// TIA Portal V15.1 export
// export: Created 2000-01-01T00:00:00.0000000Z, ExportSetting None
FUNCTION "FC_Rung" : Void   // FC42, LAD
{ S7_Optimized_Access := 'TRUE' }
   VAR_INPUT
      Local : Int;
   END_VAR
BEGIN

REGION Network 1
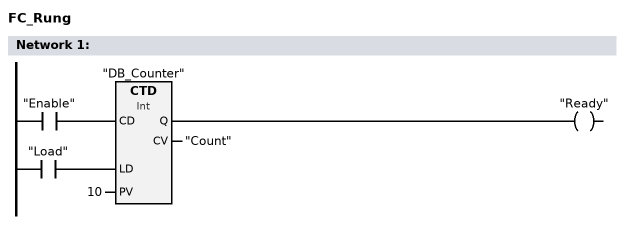
   RUNG wire#powerrail
      Contact( "Enable" )
      { S7_Templates := "value_type := Int" } "DB_Counter".CTD(ld := wire#w1, pv := 10, cv => "Count")
      Coil( "Ready" )
   END_RUNG
   RUNG wire#powerrail
      Contact( "Load" )
   END_RUNG wire#w1
   // the same network as SCL:
   "DB_Counter".CTD(CD := "Enable", LD := "Load", PV := 10, CV => "Count");
   "Ready" := "DB_Counter".Q;
END_REGION
END_FUNCTION
